Staubli VAL3: computeSPoint.pgx

public program computeSPoint(num x_nIndex, bool& x_bResult)
  local tool l_tTool
  local pointRx l_pHere
  local trsf l_trsf
  local num l_nDistance
begin
  //link(l_tTool,flange)
  //call savedata:getTool(nToolIndex,l_tTool)
  l_pHere=here(flange,world)
  l_trsf=safeTemp:sSPoint[x_nIndex].pPointRx.trsf
  l_nDistance=distance(l_pHere.trsf,l_trsf)
  if abs(l_nDistance)<5
    x_bResult=true
  else
    x_bResult=false
  endIf
end
